(* IEC 61131-3 sources: brew/plant/generated/lite/openplc/plc-power, 1 file *)

(* ---- located_vars.st ---- *)
(* Generated by plantgen from plant/plant.yaml (variant lite). Do not edit. *)
(* Analog values are raw registers: engineering value = raw / 10^scaling. *)
(* RIO I/O is at %IX100.0 / %QX100.0 / %IW100 / %QW100 (v3 and v4 alike). *)
(* PLC memory: bits from %QX0.0 (coils), words from %MW0 (holding register qw_count and up, see modbus_slave.json). *)
VAR
  PWR_MAIN_JT01_PV AT %IW100 : INT; (* Service real power (import positive), kW, x10 *)
  PWR_MAIN_JT01_ALM_HIGH AT %QX0.0 : BOOL; (* Service real power (import positive): high alarm (medium) *)
  PWR_MAIN_JT02_PV AT %IW101 : INT; (* Service reactive power, kvar, x10 *)
  PWR_MAIN_ET01_PV AT %IW102 : UINT; (* Service voltage, line to line, V, x10 *)
  PWR_MAIN_ET01_ALM_LOW AT %QX0.1 : BOOL; (* Service voltage, line to line: low alarm (medium) *)
  PWR_MAIN_IT01_PV AT %IW103 : UINT; (* Service current, phase A, A, x10 *)
  PWR_MAIN_ST01_PV AT %IW104 : UINT; (* Service frequency, Hz, x100 *)
  PWR_MAIN_JQ01_PV AT %IW105 : UINT; (* 15-minute demand (meter), kW, x10 *)
  PWR_MAIN_ZS01_PV AT %IX100.0 : BOOL; (* 52-M main breaker closed *)
  PWR_MAIN_YA01_PV AT %IX100.1 : BOOL; (* 52-M tripped on overcurrent *)
  PWR_MAIN_YA01_ALM_STATE AT %QX0.2 : BOOL; (* 52-M tripped on overcurrent: state alarm (high) *)
  PWR_MAIN_HS01_CMD AT %QX100.0 : BOOL; (* 52-M close command (0 opens) *)
  PWR_MAIN_ZS02_PV AT %IX100.2 : BOOL; (* Boiler feeder closed *)
  PWR_MAIN_ZS03_PV AT %IX100.3 : BOOL; (* Packaging feeder (PP-PKG) closed *)
  PWR_MAIN_ZS04_PV AT %IX100.4 : BOOL; (* RTU-1 feeder closed *)
  PWR_MAIN_HS02_CMD AT %QX100.1 : BOOL; (* Boiler feeder close command *)
  PWR_MAIN_HS03_CMD AT %QX100.2 : BOOL; (* Packaging feeder close command *)
  PWR_MAIN_HS04_CMD AT %QX100.3 : BOOL; (* RTU-1 feeder close command *)
  PWR_PV_JT01_PV AT %IW106 : UINT; (* PV inverter output, kW, x10 *)
  PWR_PV_JY01_PV AT %IW107 : UINT; (* PV active power limit in effect (min of site and utility), %, x10 *)
  PWR_PV_ZS01_PV AT %IX100.5 : BOOL; (* PV inverter connected (IEEE 1547) *)
  PWR_PV_HS01_CMD AT %QX100.4 : BOOL; (* PV inverter enable *)
  PWR_PV_JC01_SP AT %QW100 : UINT; (* PV site limit (plc-power), %, x10 *)
  PWR_PV_JC02_SP AT %IW108 : UINT; (* PV utility limit (DERMS through rtu-der; read only here), %, x10 *)
  PWR_BESS_JT01_PV AT %IW109 : INT; (* BESS power (discharge positive), kW, x10 *)
  PWR_BESS_EY01_PV AT %IW110 : UINT; (* BESS state of charge, %, x10 *)
  PWR_BESS_EY01_ALM_LOW AT %QX0.3 : BOOL; (* BESS state of charge: low alarm (low) *)
  PWR_BESS_ZS01_PV AT %IX100.6 : BOOL; (* BESS connected (IEEE 1547) *)
  PWR_BESS_YA01_PV AT %IX100.7 : BOOL; (* BESS PCS fault *)
  PWR_BESS_YA01_ALM_STATE AT %QX0.4 : BOOL; (* BESS PCS fault: state alarm (medium) *)
  PWR_BESS_HS01_CMD AT %QX100.5 : BOOL; (* BESS enable *)
  PWR_BESS_JC01_SP AT %QW101 : INT; (* BESS power setpoint (plc-power dispatch), kW, x10 *)
  PWR_BESS_JC02_SP AT %IW113 : INT; (* BESS utility dispatch (DERMS through rtu-der; read only here), kW, x10 *)
  PWR_BESS_TT01_PV AT %IW111 : UINT; (* BESS hottest cell temperature (BMS), degF, x10 *)
  PWR_BESS_TT01_ALM_HIGH AT %QX0.5 : BOOL; (* BESS hottest cell temperature (BMS): high alarm (medium) *)
  PWR_BESS_TT01_ALM_HIGHHIGH AT %QX0.6 : BOOL; (* BESS hottest cell temperature (BMS): highhigh alarm (high) *)
  PWR_BESS_AT01_PV AT %IW112 : UINT; (* BESS enclosure off-gas detector (electrolyte vapor; NFPA 855, UL 9540A), ppm, x1 *)
  PWR_BESS_AT01_ALM_HIGH AT %QX0.7 : BOOL; (* BESS enclosure off-gas detector (electrolyte vapor; NFPA 855, UL 9540A): high alarm (critical) *)
  PWR_GEN_JT01_PV AT %IW114 : UINT; (* Genset output, kW, x10 *)
  PWR_GEN_JT02_PV AT %IW115 : UINT; (* EP-1 emergency panel load, kW, x10 *)
  PWR_GEN_LT01_PV AT %IW116 : UINT; (* Genset fuel level, %, x10 *)
  PWR_GEN_YS01_PV AT %IX101.0 : BOOL; (* Genset running *)
  PWR_GEN_ZS01_PV AT %IX101.1 : BOOL; (* ATS on the emergency source *)
  PWR_GEN_ZS01_ALM_STATE AT %QX1.0 : BOOL; (* ATS on the emergency source: state alarm (high) *)
  PWR_GEN_ZS02_PV AT %IX101.2 : BOOL; (* Utility source available at the ATS *)
  PWR_GEN_HS01_CMD AT %QX100.6 : BOOL; (* Genset remote start (weekly exercise) *)
  PWR_GEN_KI01_PV AT %IW117 : UINT; (* ATS controller clock, minute of the local day, min, x1 *)
  PWR_GEN_KI02_PV AT %IW118 : UINT; (* ATS controller clock, local date (days since 1970-01-01), d, x1 *)
  PWR_GEN_KI03_PV AT %IW119 : UINT; (* ATS controller clock, calendar month, mo, x1 *)
  PWR_DMD_JY01_SP AT %MW0 : UINT; (* Monthly demand cap target, kW, x1 *)
  PWR_DMD_JY02_PV AT %MW1 : UINT; (* Month-to-date peak 15-minute demand, kW, x1 *)
  PWR_DMD_EY01_SP AT %MW2 : UINT; (* BESS minimum state of charge before 05:00 on brew days, %, x1 *)
  PWR_DMD_XS01_ONPEAK AT %QX1.1 : BOOL; (* SV-SGT on-peak window (weekdays 17:00-21:00) *)
  PWR_DMD_XS02_SHED AT %QX1.2 : BOOL; (* Load shed active (large feeders held open) *)
  PWR_DMD_XS03_BREWDAY AT %QX1.3 : BOOL; (* Brew day scheduled (the next 05:00 starts one; the batch engine or an operator sets it) *)
  PWR_DMD_XS04_EXERCISE AT %QX1.4 : BOOL; (* Genset exercise in progress (ATS on the genset, utility healthy) *)
  PWR_DMD_XS05_CLKOK AT %QX1.5 : BOOL; (* ATS clock trusted (in range, advancing, in step) *)
  PWR_DMD_XS05_ALM_STATE AT %QX1.6 : BOOL; (* ATS clock trusted (in range, advancing, in step): state alarm (medium) *)
END_VAR
